# EPICS autosave request: utcaApp/Db/orbit_intlk.req
$(P)$(R)IntlkEn-Sel
$(P)$(R)IntlkMinSumEn-Sel
$(P)$(R)IntlkPosEn-Sel
$(P)$(R)IntlkAngEn-Sel
$(P)$(R)IntlkLmtMinSum-SP
$(P)$(R)IntlkLmtPosMaxX-SP
$(P)$(R)IntlkLmtPosMaxY-SP
$(P)$(R)IntlkLmtAngMaxX-SP
$(P)$(R)IntlkLmtAngMaxY-SP
$(P)$(R)IntlkLmtPosMinX-SP
$(P)$(R)IntlkLmtPosMinY-SP
$(P)$(R)IntlkLmtAngMinX-SP
$(P)$(R)IntlkLmtAngMinY-SP
